FUNCTION_BLOCK FB_SimpleNcControl IMPLEMENTS I_NC_Ctrl
VAR CONSTANT
	VELO:				LREAL := 50;
END_VAR
VAR
	bEnable:			BOOL := TRUE;
	bReset:				BOOL;
	eState:				E_NC_State;
	bBusy:				BOOL;
	fbError:			FB_Error;

	
	rAxisX:				REFERENCE TO AXIS_REF;
	rAxisY:				REFERENCE TO AXIS_REF;
	rAxisZ:				REFERENCE TO AXIS_REF;
	
	fbAxisCtrlX:		FB_AxisCtrl;
	fbAxisCtrlY:		FB_AxisCtrl;
	fbAxisCtrlZ:		FB_AxisCtrl;
	
		
	fTargetX:			LREAL;
	fTargetY:			LREAL;
	fTargetZ:			LREAL;
		
	nRunState:			USINT; //0: Fall wählen; 10: nach oben, dann zum Ziel; 20: über Ziel fahren, dann senkrecht herunter //ZIEL: Gefahrenbereich umfahren
END_VAR

CASE eState OF	
	E_NC_State_INIT:
		IF __ISVALIDREF(rAxisX) AND __ISVALIDREF(rAxisY) AND __ISVALIDREF(rAxisZ) THEN			
			eState := E_NC_State_IDLE;
		END_IF

	E_NC_State_IDLE:
		;		
				
	E_NC_State_RUN:
		IF bEnable THEN
			CASE nRunState OF
				0:
					IF rAxisZ.NcToPlc.SetPos < MIN_MOVE_HEIGHT_Z AND (ABS(fTargetX - rAxisX.NcToPlc.SetPos) > 2 OR ABS(fTargetY - rAxisY.NcToPlc.SetPos) > 2) THEN
						nRunState := 10; //erst vertikal Gefahrenbereich verlassen, dann zum Ziel fahren
					ELSIF fTargetZ < MIN_MOVE_HEIGHT_Z AND (ABS(fTargetX - rAxisX.NcToPlc.SetPos) > 2 OR ABS(fTargetY - rAxisY.NcToPlc.SetPos) > 2) THEN
						nRunState := 20;
					ELSE
						nRunState := 11;
					END_IF
				
				10: //nach oben, dann zum Ziel
					fbAxisCtrlZ(stAxis := rAxisZ, eCommandIn := E_AxesCmd_MOVE_ABS, fPos := MIN_MOVE_HEIGHT_Z, fVelo := VELO);
					IF NOT fbAxisCtrlZ.bBusy THEN
						IF fbAxisCtrlZ.fbError.bError THEN
							fbError.M_Set(fbAxisCtrlZ.fbError.nErrorID, CONCAT('Achse Z: ', fbAxisCtrlZ.fbError.sErrorMsg), eState, eID := E_ErrorIDs.eAxisError, eSrc := E_ErrorSrcs.eAxisZ);
							eState := E_NC_State_ERROR;
						ELSE
							fbAxisCtrlZ(stAxis := rAxisZ, eCommandIn := E_AxesCmd_IDLE);
							nRunState := 0;
						END_IF
					END_IF
					
				11:
					fbAxisCtrlX(stAxis := rAxisX, eCommandIn := E_AxesCmd_MOVE_ABS, fPos := fTargetX, fVelo := VELO);
					fbAxisCtrlY(stAxis := rAxisY, eCommandIn := E_AxesCmd_MOVE_ABS, fPos := fTargetY, fVelo := VELO);
					fbAxisCtrlZ(stAxis := rAxisZ, eCommandIn := E_AxesCmd_MOVE_ABS, fPos := fTargetZ, fVelo := VELO);
					IF NOT fbAxisCtrlX.bBusy AND NOT fbAxisCtrlY.bBusy AND NOT fbAxisCtrlZ.bBusy THEN
						IF fbAxisCtrlX.fbError.bError THEN
							fbError.M_Set(fbAxisCtrlX.fbError.nErrorID, CONCAT('Achse X: ', fbAxisCtrlX.fbError.sErrorMsg), eState, eID := E_ErrorIDs.eAxisError, eSrc := E_ErrorSrcs.eAxisX);
							eState := E_NC_State_ERROR;
						ELSIF fbAxisCtrlY.fbError.bError THEN
							fbError.M_Set(fbAxisCtrlY.fbError.nErrorID, CONCAT('Achse Y: ', fbAxisCtrlY.fbError.sErrorMsg), eState, eID := E_ErrorIDs.eAxisError, eSrc := E_ErrorSrcs.eAxisY);
							eState := E_NC_State_ERROR;
						ELSIF fbAxisCtrlZ.fbError.bError THEN
							fbError.M_Set(fbAxisCtrlZ.fbError.nErrorID, CONCAT('Achse Z: ', fbAxisCtrlZ.fbError.sErrorMsg), eState, eID := E_ErrorIDs.eAxisError, eSrc := E_ErrorSrcs.eAxisZ);
							eState := E_NC_State_ERROR;
						ELSE
							fbAxisCtrlX(stAxis := rAxisX, eCommandIn := E_AxesCmd_IDLE);
							fbAxisCtrlY(stAxis := rAxisY, eCommandIn := E_AxesCmd_IDLE);
							fbAxisCtrlZ(stAxis := rAxisZ, eCommandIn := E_AxesCmd_IDLE);
							bBusy := FALSE;
							nRunState := 0;
							eState := E_NC_State_IDLE;
						END_IF
					END_IF
					
					
				20: //über Ziel fahren, dann senkrecht herunter
					fbAxisCtrlX(stAxis := rAxisX, eCommandIn := E_AxesCmd_MOVE_ABS, fPos := fTargetX, fVelo := VELO);
					fbAxisCtrlY(stAxis := rAxisY, eCommandIn := E_AxesCmd_MOVE_ABS, fPos := fTargetY, fVelo := VELO);
					fbAxisCtrlZ(stAxis := rAxisZ, eCommandIn := E_AxesCmd_MOVE_ABS, fPos := MIN_MOVE_HEIGHT_Z, fVelo := VELO);
					IF NOT fbAxisCtrlX.bBusy AND NOT fbAxisCtrlY.bBusy AND NOT fbAxisCtrlZ.bBusy THEN
						IF fbAxisCtrlX.fbError.bError THEN
							fbError.M_Set(fbAxisCtrlX.fbError.nErrorID, CONCAT('Achse X: ', fbAxisCtrlX.fbError.sErrorMsg), eState, eID := E_ErrorIDs.eAxisError, eSrc := E_ErrorSrcs.eAxisX);
							eState := E_NC_State_ERROR;
						ELSIF fbAxisCtrlY.fbError.bError THEN
							fbError.M_Set(fbAxisCtrlY.fbError.nErrorID, CONCAT('Achse Y: ', fbAxisCtrlY.fbError.sErrorMsg), eState, eID := E_ErrorIDs.eAxisError, eSrc := E_ErrorSrcs.eAxisY);
							eState := E_NC_State_ERROR;
						ELSIF fbAxisCtrlZ.fbError.bError THEN
							fbError.M_Set(fbAxisCtrlZ.fbError.nErrorID, CONCAT('Achse Z: ', fbAxisCtrlZ.fbError.sErrorMsg), eState, eID := E_ErrorIDs.eAxisError, eSrc := E_ErrorSrcs.eAxisZ);
							eState := E_NC_State_ERROR;
						ELSE
							fbAxisCtrlX(stAxis := rAxisX, eCommandIn := E_AxesCmd_IDLE);
							fbAxisCtrlY(stAxis := rAxisY, eCommandIn := E_AxesCmd_IDLE);
							fbAxisCtrlZ(stAxis := rAxisZ, eCommandIn := E_AxesCmd_IDLE);
							nRunState := 21;
						END_IF
					END_IF
				21:
					fbAxisCtrlZ(stAxis := rAxisZ, eCommandIn := E_AxesCmd_MOVE_ABS, fPos := fTargetZ, fVelo := VELO);
					IF NOT fbAxisCtrlZ.bBusy THEN
						IF fbAxisCtrlZ.fbError.bError THEN
							fbError.M_Set(fbAxisCtrlZ.fbError.nErrorID, CONCAT('Achse Z: ', fbAxisCtrlZ.fbError.sErrorMsg), eState, eID := E_ErrorIDs.eAxisError, eSrc := E_ErrorSrcs.eAxisZ);
							eState := E_NC_State_ERROR;
						ELSE
							fbAxisCtrlZ(stAxis := rAxisZ, eCommandIn := E_AxesCmd_IDLE);
							bBusy := FALSE;
							nRunState := 0;
							eState := E_NC_State_IDLE;
						END_IF
					END_IF
					
			END_CASE			
		ELSE
			eState := E_NC_State_ABORT;
		END_IF
		
	E_NC_State_ABORT:
		fbAxisCtrlX(stAxis := rAxisX);
		fbAxisCtrlY(stAxis := rAxisY);
		fbAxisCtrlZ(stAxis := rAxisZ);
		IF NOT fbAxisCtrlX.bBusy AND NOT fbAxisCtrlY.bBusy AND NOT fbAxisCtrlZ.bBusy THEN
			IF fbAxisCtrlX.fbError.bError THEN
				fbError.M_Set(fbAxisCtrlX.fbError.nErrorID, CONCAT('Achse X: ', fbAxisCtrlX.fbError.sErrorMsg), eState, eID := E_ErrorIDs.eAxisError, eSrc := E_ErrorSrcs.eAxisX);
				eState := E_NC_State_ERROR;
			ELSIF fbAxisCtrlY.fbError.bError THEN
				fbError.M_Set(fbAxisCtrlY.fbError.nErrorID, CONCAT('Achse Y: ', fbAxisCtrlY.fbError.sErrorMsg), eState, eID := E_ErrorIDs.eAxisError, eSrc := E_ErrorSrcs.eAxisY);
				eState := E_NC_State_ERROR;
			ELSIF fbAxisCtrlZ.fbError.bError THEN
				fbError.M_Set(fbAxisCtrlZ.fbError.nErrorID, CONCAT('Achse Z: ', fbAxisCtrlZ.fbError.sErrorMsg), eState, eID := E_ErrorIDs.eAxisError, eSrc := E_ErrorSrcs.eAxisZ);
				eState := E_NC_State_ERROR;
			ELSE
				eState := E_NC_State_IDLE;
			END_IF
		END_IF
		
	E_NC_State_ERROR:
		;
END_CASE

IF bReset THEN
	bReset := FALSE;
	fbError.M_Reset();
	IF eState = E_NC_State_ERROR THEN
		fbAxisCtrlX(stAxis := rAxisX, bReset := TRUE);
		fbAxisCtrlY(stAxis := rAxisY, bReset := TRUE);
		fbAxisCtrlZ(stAxis := rAxisZ, bReset := TRUE);
		eState := E_NC_State_IDLE;
	END_IF
END_IF

bBusy := eState <> E_NC_State_IDLE
	 AND eState <> E_NC_State_ERROR;

METHOD M_AxesReady : BOOL
VAR_INPUT
END_VAR

IF __ISVALIDREF(rAxisX) AND __ISVALIDREF(rAxisY) AND __ISVALIDREF(rAxisZ) THEN		
	rAxisX.ReadStatus();
	rAxisY.ReadStatus();
	rAxisZ.ReadStatus();
	IF rAxisX.Status.Operational AND rAxisY.Status.Operational AND rAxisZ.Status.Operational THEN
		M_AxesReady := TRUE;
	END_IF
END_IF
END_METHOD

METHOD M_AxisRef
VAR_INPUT
	rX: REFERENCE TO AXIS_REF;
	rY: REFERENCE TO AXIS_REF;
	rZ: REFERENCE TO AXIS_REF;
END_VAR

rAxisX REF= rX;
rAxisY REF= rY;
rAxisZ REF= rZ;
END_METHOD

METHOD M_CancelJob
fbAxisCtrlX(stAxis := rAxisX, eCommandIn := E_AxesCmd_IDLE);
fbAxisCtrlY(stAxis := rAxisY, eCommandIn := E_AxesCmd_IDLE);
fbAxisCtrlZ(stAxis := rAxisZ, eCommandIn := E_AxesCmd_IDLE);
eState := E_NC_State_ABORT;
END_METHOD

METHOD M_Cyclic
THIS^();

//fbAxesEnable(bEnableAxes := bEnable OR eState <> E_NC_State_IDLE, fOverride := AXES_OVERRIDE, stX := rAxisX, stY := rAxisY, stZ := rAxisZ);
fbAxisCtrlX(stAxis := rAxisX);
fbAxisCtrlY(stAxis := rAxisY);
fbAxisCtrlZ(stAxis := rAxisZ);
END_METHOD

METHOD M_NewJob
VAR_INPUT
	fTargetPosX	: LREAL;
	fTargetPosY	: LREAL;
	fTargetPosZ	: LREAL;
END_VAR
IF M_AxesReady() THEN
	IF eState = E_NC_State_IDLE THEN
		fTargetX := fTargetPosX;
		fTargetY := fTargetPosY;
		fTargetZ := fTargetPosZ;
		eState := E_NC_State_RUN;
		nRunState := 0;
		fbError.M_Reset();
	ELSIF eState = E_NC_State_RUN AND (fTargetX <> fTargetPosX OR fTargetY <> fTargetPosY OR fTargetZ <> fTargetPosZ) THEN	
		M_CancelJob();
	END_IF
ELSE
	fbError.M_Set(1, 'Achsen sind nicht bereit!', eState, eID := E_ErrorIDs.eAxesNotReady, eSrc := E_ErrorSrcs.eAxisCtrlPtp);
END_IF
END_METHOD


PROPERTY P_Busy : BOOL
GET
P_Busy := bBusy;
END_GET
END_PROPERTY

PROPERTY P_Enable : BOOL
SET
bEnable := P_Enable;
END_SET
END_PROPERTY

PROPERTY P_ErrID : UDINT
GET
P_ErrID := fbError.nErrorID;
END_GET
END_PROPERTY

PROPERTY P_ErrMsg : STRING
GET
P_ErrMsg := fbError.sErrorMsg;
END_GET
END_PROPERTY

PROPERTY P_Error : BOOL
GET
P_Error := fbError.bError;
END_GET
END_PROPERTY


PROPERTY P_Reset : BOOL
SET
bReset := P_Reset;
END_SET
END_PROPERTY

END_FUNCTION_BLOCK

(* stored: Version 1.1.0.1, ProductVersion 3.1.4024.9
   POU FB_SimpleNcControl: Id {c236e9e8-0263-42e9-82d1-aa06de294b98}, SpecialFunc None
   Method M_AxesReady: Id {c8a10f5e-82d0-4b35-9242-c490062659ae}
   Method M_AxisRef: Id {dcca78ad-e6bb-4717-a84e-0d5c88ba4d6b}
   Method M_CancelJob: Id {3fe2cf29-9c01-4b25-89e9-4a8027f76695}
   Method M_Cyclic: Id {7e4f8fa1-fcb0-42e3-9b6d-09a9858a4de8}
   Method M_NewJob: Id {ca4ee68f-6e3a-4e4e-aeed-8d6a5345539a}
   Property P_Busy: Id {3887cb1c-0457-4933-847d-51378cb220ed}
   Get Get: Id {b41cbe41-4a13-44ba-b768-1f234dbcf707}
   Property P_Enable: Id {f7e7b5bb-ba54-40e7-b06c-2e2add145769}
   Set Set: Id {13ccb6e4-22e3-4365-b80f-9e50af8a9003}
   Property P_ErrID: Id {876b6736-0bf5-4b8e-a55c-eab4c330f51e}
   Get Get: Id {b1fa7b41-37cd-4407-8f74-cf35577c637f}
   Property P_ErrMsg: Id {7f637b45-e7fe-41a6-aadc-a61535c0c11c}
   Get Get: Id {e2bdb9f5-f7df-4188-8b95-e3f687ff2583}
   Property P_Error: Id {aa27c985-30ac-4631-b09f-6387107b74f7}
   Get Get: Id {28a120ad-575a-43b9-b0e1-bd7f0d410949}
   Property P_Reset: Id {979f83c8-5916-4d66-ac03-6e9589efbfd8}
   Set Set: Id {1da12ba2-b9e3-441e-9334-397cd7abb3ca} *)
